(* IEC 61131-3 sources: plc-cip-batch-control/plc/prog, 5 files *)

(* ---- PRG_Alarms.st ---- *)
(*
    PRG_Alarms.st: the alarm list.

    Twelve points, each with a priority and an on-delay chosen so that the
    operator is not told about things that resolve themselves. ISA-18.2's first
    rule is that every alarm must require a response; a low chemical level that
    clears in two seconds does not.

    First-out is captured and held until the list goes quiet, so the record
    says which condition started the trip rather than which one is loudest by
    the time anyone looks.
*)

PROGRAM PRG_Alarms
VAR
    fbSafety        : FB_Alarm;
    fbSupplyPump    : FB_Alarm;
    fbReturnPump    : FB_Alarm;
    fbLevelLow      : FB_Alarm;
    fbCausticLow    : FB_Alarm;
    fbAcidLow       : FB_Alarm;
    fbTempLow       : FB_Alarm;
    fbFlowLow       : FB_Alarm;
    fbCircuitBusy   : FB_Alarm;
    fbPhaseTimeout  : FB_Alarm;
    fbNotClean      : FB_Alarm;
    fbNoSteam       : FB_Alarm;
    fbCondSensor    : FB_Alarm;
    i               : INT;
    xAnyLatched     : BOOL;
    xCirculating    : BOOL;
END_VAR

xCirculating := gxPhaseExecute AND (gPhaseStep = PS_CIRCULATE);

fbSafety(xCondition := gxSafetyTrip,
         iPriority  := 1,
         xAck       := xCmdAckAlarms,
         rNowS      := grPlcTimeS,
         stAlarm    := gAlarms[C_ALM_SAFETY]);

fbSupplyPump(xCondition := xSupplyPumpFault OR (xSupplyPumpRun AND NOT xSupplyPumpRunning),
             iPriority  := 1,
             tOnDelay   := T#5s,
             xAck       := xCmdAckAlarms,
             rNowS      := grPlcTimeS,
             stAlarm    := gAlarms[C_ALM_SUPPLY_PUMP]);

fbReturnPump(xCondition := xReturnPumpFault OR (xReturnPumpRun AND NOT xReturnPumpRunning),
             iPriority  := 2,
             tOnDelay   := T#5s,
             xAck       := xCmdAckAlarms,
             rNowS      := grPlcTimeS,
             stAlarm    := gAlarms[C_ALM_RETURN_PUMP]);

fbLevelLow(xCondition := (rLevelBalanceTankPct < C_LEVEL_TRIP_PCT) AND (gUnitState <> UST_IDLE),
           iPriority  := 2,
           tOnDelay   := T#3s,
           xAck       := xCmdAckAlarms,
           rNowS      := grPlcTimeS,
           stAlarm    := gAlarms[C_ALM_LEVEL_LOW]);

fbCausticLow(xCondition := rLevelCausticPct < C_CHEM_LEVEL_MIN,
             iPriority  := 3,
             tOnDelay   := T#10s,
             xAck       := xCmdAckAlarms,
             rNowS      := grPlcTimeS,
             stAlarm    := gAlarms[C_ALM_CAUSTIC_LOW]);

fbAcidLow(xCondition := rLevelAcidPct < C_CHEM_LEVEL_MIN,
          iPriority  := 3,
          tOnDelay   := T#10s,
          xAck       := xCmdAckAlarms,
          rNowS      := grPlcTimeS,
          stAlarm    := gAlarms[C_ALM_ACID_LOW]);

(* Twelve minutes: a cold circuit and a 1200 litre balance tank take about
   eight to come up to a wash temperature, so anything shorter alarms on every
   normal start. It still catches a steam valve that never opened. *)
fbTempLow(xCondition := xCirculating AND gPhaseParams.xHeat
                        AND (rTempReturnC < gPhaseParams.rTempMin),
          iPriority  := 2,
          tOnDelay   := T#12m,
          xAck       := xCmdAckAlarms,
          rNowS      := grPlcTimeS,
          stAlarm    := gAlarms[C_ALM_TEMP_LOW]);

fbFlowLow(xCondition := xCirculating AND (rFlowSupplyM3h < gPhaseParams.rFlowMin),
          iPriority  := 2,
          tOnDelay   := T#30s,
          xAck       := xCmdAckAlarms,
          rNowS      := grPlcTimeS,
          stAlarm    := gAlarms[C_ALM_FLOW_LOW]);

fbCircuitBusy(xCondition := (NOT xCircuitAvailable) AND (gUnitState <> UST_IDLE),
              iPriority  := 2,
              tOnDelay   := T#3s,
              xAck       := xCmdAckAlarms,
              rNowS      := grPlcTimeS,
              stAlarm    := gAlarms[C_ALM_CIRCUIT_BUSY]);

fbPhaseTimeout(xCondition := (gFailCode = FC_PHASE_TIMEOUT) OR (gFailCode = FC_CHARGE_TIMEOUT)
                             OR (gFailCode = FC_TEMP_TIMEOUT),
               iPriority  := 1,
               xAck       := xCmdAckAlarms,
               rNowS      := grPlcTimeS,
               stAlarm    := gAlarms[C_ALM_PHASE_TIMEOUT]);

fbNotClean(xCondition := gFailCode = FC_RINSE_NOT_CLEAN,
           iPriority  := 1,
           xAck       := xCmdAckAlarms,
           rNowS      := grPlcTimeS,
           stAlarm    := gAlarms[C_ALM_NOT_CLEAN]);

fbNoSteam(xCondition := (NOT xSteamAvailable) AND gPhaseParams.xHeat AND gxPhaseExecute,
          iPriority  := 3,
          tOnDelay   := T#10s,
          xAck       := xCmdAckAlarms,
          rNowS      := grPlcTimeS,
          stAlarm    := gAlarms[C_ALM_NO_STEAM]);

fbCondSensor(xCondition := gxCondSensorFault,
             iPriority  := 1,
             xAck       := xCmdAckAlarms,
             rNowS      := grPlcTimeS,
             stAlarm    := gAlarms[C_ALM_COND_SENSOR]);

(* ---- summary ---------------------------------------------------------- *)
giActiveAlarms := 0;
gxAlarmP1Active := FALSE;
xAnyLatched := FALSE;
xHmiAlarmHorn := FALSE;

FOR i := 1 TO C_ALARM_COUNT DO
    IF gAlarms[i].xLatched THEN
        xAnyLatched := TRUE;
        giActiveAlarms := giActiveAlarms + 1;
        IF gAlarms[i].xActive AND (gAlarms[i].iPriority = 1) THEN
            gxAlarmP1Active := TRUE;
        END_IF
        IF NOT gAlarms[i].xAcked THEN
            xHmiAlarmHorn := TRUE;
        END_IF
        IF giFirstOut = 0 THEN
            giFirstOut := i;
        END_IF
    END_IF
END_FOR

IF NOT xAnyLatched THEN
    giFirstOut := 0;
END_IF

(* Acknowledge is momentary too and this is the last program that reads it. *)
xCmdAckAlarms := FALSE;

END_PROGRAM

(* ---- PRG_Control.st ---- *)
(*
    PRG_Control.st: the only program that writes to the field outputs.

    It takes the demand PRG_Sequence produced, applies the permissives
    PRG_Safety produced and drives the valve matrix, the two motor starters
    and the two closed loops. Because it is the single writer, the question
    "what could possibly open the steam valve?" has exactly one answer.

    Loops:
      flow  -> supply pump speed, PI. Slow, because the pump is a VSD against
               a fixed circuit resistance and there is nothing to gain from
               being quick.
      temperature -> steam valve, PI on the supply temperature. Tuned soft:
               the plate pack has a couple of seconds of transport delay and
               the balance tank behind it is a 1200 litre integrator.
*)

PROGRAM PRG_Control
VAR
    fbFlowPid       : FB_Pid;
    fbTempPid       : FB_Pid;
    fbSupplyLimit   : FB_Pid;
    fbSupplyPump    : FB_Pump;
    fbReturnPump    : FB_Pump;
    xRunSupply      : BOOL;
    xRunReturn      : BOOL;
    xHeatDemand     : BOOL;
    xDoseDemand     : BOOL;
END_VAR

(* ---- interlocked demands --------------------------------------------- *)
xRunSupply  := gDemand.xSupplyPump AND gxPermitRun;
xRunReturn  := gDemand.xReturnPump AND gxPermitRun;
xHeatDemand := gDemand.xHeat AND gxPermitHeat;
xDoseDemand := gDemand.xDose AND gxPermitDose;

(* ---- motor starters --------------------------------------------------- *)
fbSupplyPump(xStart       := xRunSupply,
             xInterlockOk := gxPermitRun,
             xRunFeedback := xSupplyPumpRunning,
             xFault       := xSupplyPumpFault,
             xReset       := xCmdReset);

fbReturnPump(xStart       := xRunReturn,
             xInterlockOk := gxPermitRun,
             xRunFeedback := xReturnPumpRunning,
             xFault       := xReturnPumpFault,
             xReset       := xCmdReset);

xSupplyPumpRun := fbSupplyPump.xRun;
xReturnPumpRun := fbReturnPump.xRun;

(* ---- flow loop -------------------------------------------------------- *)
fbFlowPid(xEnable := fbSupplyPump.xRun,
          rPv     := rFlowSupplyM3h,
          rSp     := gDemand.rFlowSp,
          rKp     := 3.0,
          rTi     := 8.0,
          rOutMin := C_PUMP_SPEED_MIN,
          rOutMax := C_PUMP_SPEED_MAX,
          rCycleS := C_CYCLE_S);

IF fbSupplyPump.xRun THEN
    rSupplyPumpSpeedPct := fbFlowPid.rOut;
ELSE
    rSupplyPumpSpeedPct := 0.0;
END_IF

(* ---- temperature loop -------------------------------------------------- *)
(* The controlled variable is the return temperature, not the supply. The
   recipe specifies a temperature at the soil and the coldest point of the
   circuit is the one that has to reach it; controlling the supply instead
   throttles the steam as soon as one pass through the plate pack looks hot
   enough and the loop then takes three times as long to bring the balance
   tank up.

   Tuning is lambda tuning for an integrator with dead time: the circuit holds
   450 litres, so at 18 m3/h a change at the plate pack takes about 90 seconds
   to reach the return element. Kp 5 %/K, Ti 600 s. *)
fbTempPid(xEnable := xHeatDemand,
          rPv     := rTempReturnC,
          rSp     := gDemand.rTempSp,
          rKp     := 5.0,
          rTi     := 600.0,
          rOutMin := 0.0,
          rOutMax := 100.0,
          rCycleS := C_CYCLE_S);

(* Override: a proportional-only high limit on the plate-pack outlet, low
   selected against the main loop. Proportional only on purpose, because an
   integrator on the losing half of a selector winds up. *)
fbSupplyLimit(xEnable := xHeatDemand,
              rPv     := rTempSupplyC,
              rSp     := C_SUPPLY_TEMP_LIMIT,
              rKp     := 25.0,
              rTi     := 0.0,
              rOutMin := 0.0,
              rOutMax := 100.0,
              rCycleS := C_CYCLE_S);

xSteamIsolation := xHeatDemand;
IF xHeatDemand THEN
    rSteamValvePct := MIN(fbTempPid.rOut, fbSupplyLimit.rOut);
ELSE
    rSteamValvePct := 0.0;
END_IF

(* ---- valve matrix ----------------------------------------------------- *)
(* Source selection. Only one inlet is ever open and the fill valve gates
   the whole group so a phase can hold its line-up without taking liquid. *)
xV01FreshWater     := gDemand.xFillValve AND (gDemand.eSource = SRC_FRESH);
xV02RecoveredWater := gDemand.xFillValve AND (gDemand.eSource = SRC_RECOVERED);
xV11CausticSupply  := gDemand.xFillValve AND (gDemand.eSource = SRC_CAUSTIC);
xV12AcidSupply     := gDemand.xFillValve AND (gDemand.eSource = SRC_ACID);

(* Dosing is concentrate trim on top of whatever the tank already holds, so it
   is gated on the phase's dose demand rather than on the fill valve. *)
xV03CausticDose    := xDoseDemand AND (gDemand.eSource = SRC_CAUSTIC);
xV04AcidDose       := xDoseDemand AND (gDemand.eSource = SRC_ACID);

xV08ReturnToCaustic := FALSE;
xV10ReturnToAcid := FALSE;

(* Return destination. Exactly one of these is open whenever the return pump
   is running, so the circuit always has somewhere to discharge. *)
xV06ReturnToDrain    := FALSE;
xV07ReturnToBalance  := FALSE;
xV09ReturnToRecovery := FALSE;

CASE gDemand.eReturn OF
    RET_DRAIN:
        xV06ReturnToDrain := TRUE;
    RET_RECOVERY:
        xV09ReturnToRecovery := TRUE;
    RET_CAUSTIC:
        xV08ReturnToCaustic := TRUE;
    RET_ACID:
        xV10ReturnToAcid := TRUE;
    RET_BALANCE:
        xV07ReturnToBalance := TRUE;
END_CASE

xV05SupplyToCircuit := fbSupplyPump.xRun;

END_PROGRAM

(* ---- PRG_Kpi.st ---- *)
(*
    PRG_Kpi.st: consumption totals, the batch record and the SCADA image.

    Everything here is computed from instruments the skid actually has: the
    make-up flow meter, the supply flow meter, the two temperature elements
    either side of the heat exchanger and the dosing pump run time. Nothing
    is inferred from the model, so the same code would produce the same batch
    record on real hardware.

    Steam energy is the enthalpy the water gained across the plate pack:

        kW = m3/h * 1000 / 3600 [kg/s] * 4.19 [kJ/kg.K] * (Tsupply - Ttank) [K]

    which under-reports the boiler's fuel by the efficiency of the pack and
    the condensate return. It is the number the site can act on and it is
    the one the utility meter can be reconciled against.
*)

PROGRAM PRG_Kpi
VAR
    fbFresh         : FB_Totaliser;
    fbRecovered     : FB_Totaliser;
    fbEffluent      : FB_Totaliser;
    fbCaustic       : FB_Totaliser;
    fbAcid          : FB_Totaliser;
    fbEnergy        : FB_Totaliser;
    rEnergyKW       : REAL;
    rSnapWater      : REAL;
    rSnapChem       : REAL;
    rSnapEnergy     : REAL;
    i               : INT;
    xAllPass        : BOOL;
    xFinalRinseOk   : BOOL;
    xUnitActive     : BOOL;
END_VAR

xUnitActive := (gUnitState <> UST_IDLE)
               AND (gUnitState <> UST_COMPLETE)
               AND (gUnitState <> UST_ABORTED);

(* ---- instantaneous steam duty ---------------------------------------- *)
IF xSteamIsolation AND (rTempSupplyC > rTempBalanceTankC) THEN
    rEnergyKW := rFlowSupplyM3h * 1000.0 / 3600.0 * 4.19 * (rTempSupplyC - rTempBalanceTankC);
ELSE
    rEnergyKW := 0.0;
END_IF

(* ---- totalisers, all reset together at the start of a batch ------------
    Each is gated on the line-up rather than on a valve command. That
    distinction matters more than it looks.

    Make-up is bang-bang level control on a break tank, so V01 and V02 toggle
    every scan or two. The flow transmitter is read at the top of the scan and
    therefore reports the previous scan's flow, so gating the totaliser on the
    valve command aliases the two signals: on the scans the valve is open the
    meter is still reporting the scan it was shut, so the total comes out
    about a fifth low. The source selection only changes at a phase boundary
    and the meter reads zero when the valve is shut in any case. Gating on
    the source and letting the low-flow cut-off reject the noise measures
    what actually went through the meter.
*)
fbFresh(xEnable := gDemand.eSource = SRC_FRESH,
        rRatePerHour := rFlowMakeupM3h * 1000.0,
        rCutOff := 50.0,
        rCycleS := C_CYCLE_S,
        xReset := gxCycleReset);

fbRecovered(xEnable := gDemand.eSource = SRC_RECOVERED,
            rRatePerHour := rFlowMakeupM3h * 1000.0,
            rCutOff := 50.0,
            rCycleS := C_CYCLE_S,
            xReset := gxCycleReset);

fbEffluent(xEnable := xV06ReturnToDrain,
           rRatePerHour := rFlowSupplyM3h * 1000.0,
           rCutOff := 50.0,
           rCycleS := C_CYCLE_S,
           xReset := gxCycleReset);

fbCaustic(xEnable := xV03CausticDose,
          rRatePerHour := C_CAUSTIC_DOSE_LPM * 60.0,
          rCycleS := C_CYCLE_S,
          xReset := gxCycleReset);

fbAcid(xEnable := xV04AcidDose,
       rRatePerHour := C_ACID_DOSE_LPM * 60.0,
       rCycleS := C_CYCLE_S,
       xReset := gxCycleReset);

fbEnergy(xEnable := xSteamIsolation,
         rRatePerHour := rEnergyKW,
         rCycleS := C_CYCLE_S,
         xReset := gxCycleReset);

gKpi.rFreshWaterL     := fbFresh.rTotal;
gKpi.rRecoveredWaterL := fbRecovered.rTotal;
gKpi.rEffluentL       := fbEffluent.rTotal;
gKpi.rCausticL        := fbCaustic.rTotal;
gKpi.rAcidL           := fbAcid.rTotal;
gKpi.rEnergyKWh       := fbEnergy.rTotal;

IF gxCycleReset THEN
    grCycleElapsedS := 0.0;
    gKpi.xVerifiedClean := FALSE;
    rSnapWater := 0.0;
    rSnapChem := 0.0;
    rSnapEnergy := 0.0;
END_IF

IF xUnitActive THEN
    grCycleElapsedS := grCycleElapsedS + C_CYCLE_S;
END_IF
gKpi.rCycleTimeS := grCycleElapsedS;

(* ---- per-phase consumption, by difference ----------------------------- *)
IF gxPhaseStartPulse THEN
    rSnapWater  := fbFresh.rTotal + fbRecovered.rTotal;
    rSnapChem   := fbCaustic.rTotal + fbAcid.rTotal;
    rSnapEnergy := fbEnergy.rTotal;
END_IF

IF gxPhaseEndPulse AND (giPhaseIndex >= 1) AND (giPhaseIndex <= C_PHASE_COUNT) THEN
    gResults[giPhaseIndex].rWaterL := fbFresh.rTotal + fbRecovered.rTotal - rSnapWater;
    gResults[giPhaseIndex].rChemL := fbCaustic.rTotal + fbAcid.rTotal - rSnapChem;
    gResults[giPhaseIndex].rEnergyKWh := fbEnergy.rTotal - rSnapEnergy;
END_IF

(* ---- release criteria -------------------------------------------------- *)
(* A batch is only released if every phase that ran met its own criteria and
   the final rinse came back as clean as the water going in. A fixed-time
   recipe can complete without satisfying the second test and that is the
   whole argument for the adaptive one. *)
xAllPass := TRUE;
FOR i := 1 TO C_PHASE_COUNT DO
    IF gResults[i].xExecuted AND NOT gResults[i].xPass THEN
        xAllPass := FALSE;
    END_IF
END_FOR

xFinalRinseOk := gResults[5].xExecuted
                 AND gResults[5].xPass
                 AND (gResults[5].rEndConductivity <= gRecipe.rRinseEndCond);

IF gUnitState = UST_COMPLETE THEN
    gKpi.xVerifiedClean := xAllPass AND xFinalRinseOk;
END_IF

(* ---- SCADA image ------------------------------------------------------- *)
iHmiUnitState        := TO_INT(gUnitState);
iHmiPhase            := TO_INT(gPhase);
iHmiPhaseStep        := TO_INT(gPhaseStep);
iHmiFailCode         := TO_INT(gFailCode);
iHmiActiveAlarms     := giActiveAlarms;
iHmiFirstOutAlarm    := giFirstOut;
iHmiBatchId          := giBatchId;

rHmiFreshWaterL      := gKpi.rFreshWaterL;
rHmiRecoveredWaterL  := gKpi.rRecoveredWaterL;
rHmiEffluentL        := gKpi.rEffluentL;
rHmiCausticL         := gKpi.rCausticL;
rHmiAcidL            := gKpi.rAcidL;
rHmiEnergyKWh        := gKpi.rEnergyKWh;
rHmiCycleTimeS       := gKpi.rCycleTimeS;
rHmiPhaseElapsedS    := grPhaseElapsedS;
rHmiHoldAchievedS    := grHoldAchievedS;
rHmiConcentrationPct := grConcentrationPct;

xHmiVerifiedClean    := gKpi.xVerifiedClean;
xHmiCycleComplete    := gUnitState = UST_COMPLETE;
xHmiCycleAborted     := gUnitState = UST_ABORTED;
xHmiHeating          := xSteamIsolation;

END_PROGRAM

(* ---- PRG_Safety.st ---- *)
(*
    PRG_Safety.st: interlocks and permissives. First program in the task, so
    every other program sees a permit that was evaluated against this scan's
    inputs rather than the previous one's.

    Nothing here is a substitute for the hard-wired safety circuit. The E-stop
    drops the contactors and the steam solenoid directly; xSafetyOk is only the
    controller's view of that circuit, used to sequence a clean shutdown.

    Two interlocks earn their place:

      * no steam without proven flow. A steam-heated plate pack with no flow
        through it will boil the film against the plate, bake the soil on and
        eventually damage the gaskets.
      * no dosing without a running supply pump and a source that has stock in
        it, so concentrate cannot sit undiluted in the balance tank.
*)

PROGRAM PRG_Safety
VAR CONSTANT
    C_MIN_FLOW_HEAT : REAL := 8.0;      (* m3/h before steam may be admitted *)
    C_DRY_RUN_FLOW  : REAL := 2.0;      (* m3/h with the pump running is a dry run *)
END_VAR
VAR
    fbDryRun        : TON;
    fbCircuitLost   : TON;
    xChemStockOk    : BOOL;
END_VAR

grPlcTimeS := grPlcTimeS + C_CYCLE_S;

(* A running pump moving nothing is either dry or dead-headed. Either way it
   destroys the seal in minutes, so it is a latch-free hard stop. *)
fbDryRun(IN := xSupplyPumpRunning AND (rFlowSupplyM3h < C_DRY_RUN_FLOW), PT := T#20s);

fbCircuitLost(IN := NOT xCircuitAvailable, PT := T#3s);

gxSafetyTrip := (NOT xSafetyOk)
                OR xBalanceTankLowLow
                OR fbDryRun.Q
                OR (gUnitState <> UST_IDLE AND fbCircuitLost.Q);

gxPermitRun := xSafetyOk
               AND (NOT xBalanceTankLowLow)
               AND (NOT fbDryRun.Q)
               AND xCircuitAvailable
               AND (rLevelBalanceTankPct > C_LEVEL_TRIP_PCT);

gxPermitHeat := gxPermitRun
                AND xSteamAvailable
                AND xSupplyPumpRunning
                AND (rFlowSupplyM3h >= C_MIN_FLOW_HEAT);

(* Only the tank the current phase is drawing from has to have stock. *)
CASE gDemand.eSource OF
    SRC_CAUSTIC:
        xChemStockOk := rLevelCausticPct > C_CHEM_LEVEL_MIN;
    SRC_ACID:
        xChemStockOk := rLevelAcidPct > C_CHEM_LEVEL_MIN;
ELSE
    xChemStockOk := TRUE;
END_CASE

gxPermitDose := gxPermitRun AND xSupplyPumpRunning AND xChemStockOk;

END_PROGRAM

(* ---- PRG_Sequence.st ---- *)
(*
    PRG_Sequence.st: the ISA-88 unit procedure.

    This program owns the unit state machine and turns the recipe into phase
    parameters. It does not touch a single output. It produces a demand;
    PRG_Control decides whether the interlocks let that demand reach the
    field. Keeping the two apart is what makes the sequence readable and the
    interlocks auditable.

    Phase order is fixed; the recipe chooses which phases are in it:

        PRE_RINSE -> CAUSTIC -> INTERMEDIATE RINSE -> [ACID] ->
        FINAL RINSE -> [SANITISE] -> COMPLETE
*)

(*
    How long a rinse must run before its conductivity endpoint means anything.

    The return element sits downstream of the whole circuit, so a rinse that
    stops after twenty seconds has only measured the water that was already in
    the pipe. The floor is one and a half circuit turnovers at the recipe flow
    (135 seconds for a 450 litre circuit at 18 m3/h) or the recipe's own
    minimum, whichever is longer.
*)
FUNCTION RinseBlankTime : TIME
VAR_INPUT
    tFloor      : TIME;
    rFlowSpM3h  : REAL;
END_VAR
VAR
    rFlowLps    : REAL;
    rTurnoverS  : REAL;
END_VAR

rFlowLps := MAX(rFlowSpM3h, 1.0) * 1000.0 / 3600.0;
rTurnoverS := C_RINSE_TURNOVERS * C_CIRCUIT_VOLUME_L / rFlowLps;
RinseBlankTime := SecondsToTime(MAX(TimeToSeconds(tFloor), rTurnoverS));

END_FUNCTION

FUNCTION NextPhase : E_Phase
VAR_INPUT
    eCurrent     : E_Phase;
    xUseAcid     : BOOL;
    xUseSanitise : BOOL;
END_VAR

CASE eCurrent OF
    PH_IDLE:
        NextPhase := PH_PRE_RINSE;
    PH_PRE_RINSE:
        NextPhase := PH_CAUSTIC_WASH;
    PH_CAUSTIC_WASH:
        NextPhase := PH_INTERMEDIATE_RINSE;
    PH_INTERMEDIATE_RINSE:
        IF xUseAcid THEN
            NextPhase := PH_ACID_WASH;
        ELSE
            NextPhase := PH_FINAL_RINSE;
        END_IF
    PH_ACID_WASH:
        NextPhase := PH_FINAL_RINSE;
    PH_FINAL_RINSE:
        IF xUseSanitise THEN
            NextPhase := PH_SANITISE;
        ELSE
            NextPhase := PH_COMPLETE;
        END_IF
    PH_SANITISE:
        NextPhase := PH_COMPLETE;
ELSE
    NextPhase := PH_COMPLETE;
END_CASE

END_FUNCTION

PROGRAM PRG_Sequence
VAR
    fbUnit          : FB_UnitStateMachine;
    fbPhase         : FB_CipPhase;
    iPhaseIndex     : INT;
    iResultIndex    : INT;
    xReadyToStart   : BOOL;
    xProcComplete   : BOOL;
    xProcFailed     : BOOL;
    xPhaseGap       : BOOL;     (* one scan between phases, re-arms the engine *)
    xPhaseActive    : BOOL;     (* running or held: the engine keeps its state *)
    xExecutePhase   : BOOL;     (* running: accumulators and alarms advance *)
    ePrevPhase      : E_Phase;
END_VAR

(* ---------------------------------------------------------------------- *)
(* 1. Unit state machine                                                    *)
(* ---------------------------------------------------------------------- *)
xReadyToStart := (NOT gxSafetyTrip) AND xCircuitAvailable AND (NOT gxAlarmP1Active);

fbUnit(xStart              := xCmdStart,
       xHold               := xCmdHold,
       xRestart            := xCmdRestart,
       xAbort              := xCmdAbort,
       xReset              := xCmdReset,
       xReadyToStart       := xReadyToStart,
       xProcedureComplete  := xProcComplete,
       xProcedureFailed    := xProcFailed,
       xSafetyTrip         := gxSafetyTrip);

gUnitState := fbUnit.eState;

(* ---------------------------------------------------------------------- *)
(* 2. Start of batch                                                        *)
(* ---------------------------------------------------------------------- *)
gxCycleReset := FALSE;
IF fbUnit.xStartPulse THEN
    giBatchId := giBatchId + 1;
    gPhase := PH_PRE_RINSE;
    gFailCode := FC_NONE;
    xProcComplete := FALSE;
    xProcFailed := FALSE;
    xPhaseGap := FALSE;
    gxCycleReset := TRUE;
    gxCondSensorFault := FALSE;
    gxCondProven := FALSE;
    FOR iPhaseIndex := 1 TO C_PHASE_COUNT DO
        gResults[iPhaseIndex].ePhase := PH_IDLE;
        gResults[iPhaseIndex].xExecuted := FALSE;
        gResults[iPhaseIndex].xPass := FALSE;
        gResults[iPhaseIndex].eFail := FC_NONE;
        gResults[iPhaseIndex].rDurationS := 0.0;
        gResults[iPhaseIndex].rHoldAchievedS := 0.0;
        gResults[iPhaseIndex].rWaterL := 0.0;
        gResults[iPhaseIndex].rChemL := 0.0;
        gResults[iPhaseIndex].rEnergyKWh := 0.0;
    END_FOR
END_IF

IF fbUnit.eState = UST_IDLE THEN
    gPhase := PH_IDLE;
    gFailCode := FC_NONE;
END_IF

(* ---------------------------------------------------------------------- *)
(* 3. Phase parameters from the recipe                                      *)
(* ---------------------------------------------------------------------- *)
gPhaseParams.rFlowSp  := gRecipe.rFlowSp;
gPhaseParams.rFlowMin := gRecipe.rFlowMin;
gPhaseParams.tMaxPhase := gRecipe.tPhaseMax;
gPhaseParams.tMinPhase := T#30s;
gPhaseParams.xAdaptiveEnd := FALSE;
gPhaseParams.rEndConductivity := gRecipe.rRinseEndCond;
gPhaseParams.rConcSp := 0.0;
gPhaseParams.rConcMin := 0.0;
gPhaseParams.rConcMax := 0.0;
gPhaseParams.rTempSp := 0.0;
gPhaseParams.rTempMin := 0.0;
gPhaseParams.xHeat := FALSE;
gPhaseParams.xDose := FALSE;
gPhaseParams.xRecirculate := FALSE;

CASE gPhase OF

    PH_PRE_RINSE:
        (* Recovered final-rinse water if there is any, mains if not. This one
           line is most of the water saving: the pre-rinse is the biggest
           single-pass consumer in the cycle. *)
        IF rLevelRecoveryPct > 25.0 THEN
            gPhaseParams.eSource := SRC_RECOVERED;
        ELSE
            gPhaseParams.eSource := SRC_FRESH;
        END_IF
        gPhaseParams.eReturn := RET_DRAIN;
        gPhaseParams.tHold := gRecipe.tPreRinse;
        gPhaseParams.tMinPhase := RinseBlankTime(gRecipe.tRinseMin, gRecipe.rFlowSp);
        gPhaseParams.tRecover := T#20s;
        gPhaseParams.tMaxPhase := gRecipe.tRinseMax;
        gPhaseParams.xAdaptiveEnd := gRecipe.xAdaptive;
        (* Gross soil removal: a looser endpoint than the final rinse. *)
        gPhaseParams.rEndConductivity := gRecipe.rRinseEndCond * 3.0;

    PH_CAUSTIC_WASH:
        gPhaseParams.eSource := SRC_CAUSTIC;
        gPhaseParams.eReturn := RET_CAUSTIC;
        gPhaseParams.xRecirculate := TRUE;
        gPhaseParams.rTempSp := gRecipe.rCausticTempSp;
        gPhaseParams.rTempMin := gRecipe.rCausticTempMin;
        gPhaseParams.xHeat := TRUE;
        gPhaseParams.rConcSp := gRecipe.rCausticConcSp;
        gPhaseParams.rConcMin := gRecipe.rCausticConcSp - 0.25;
        gPhaseParams.rConcMax := gRecipe.rCausticConcSp + 0.50;
        gPhaseParams.xDose := TRUE;
        gPhaseParams.tHold := gRecipe.tCausticHold;
        gPhaseParams.tMinPhase := T#1m;
        gPhaseParams.tRecover := T#180s;

    PH_INTERMEDIATE_RINSE:
        gPhaseParams.eSource := SRC_FRESH;
        gPhaseParams.eReturn := RET_DRAIN;
        gPhaseParams.tHold := gRecipe.tIntRinse;
        gPhaseParams.tMinPhase := RinseBlankTime(gRecipe.tRinseMin, gRecipe.rFlowSp);
        gPhaseParams.tRecover := T#20s;
        gPhaseParams.tMaxPhase := gRecipe.tRinseMax;
        gPhaseParams.xAdaptiveEnd := gRecipe.xAdaptive;
        gPhaseParams.rEndConductivity := gRecipe.rRinseEndCond * 2.0;

    PH_ACID_WASH:
        gPhaseParams.eSource := SRC_ACID;
        gPhaseParams.eReturn := RET_ACID;
        gPhaseParams.xRecirculate := TRUE;
        gPhaseParams.rTempSp := gRecipe.rAcidTempSp;
        gPhaseParams.rTempMin := gRecipe.rAcidTempMin;
        gPhaseParams.xHeat := TRUE;
        gPhaseParams.rConcSp := gRecipe.rAcidConcSp;
        gPhaseParams.rConcMin := gRecipe.rAcidConcSp - 0.15;
        gPhaseParams.rConcMax := gRecipe.rAcidConcSp + 0.35;
        gPhaseParams.xDose := TRUE;
        gPhaseParams.tHold := gRecipe.tAcidHold;
        gPhaseParams.tMinPhase := T#1m;
        gPhaseParams.tRecover := T#180s;

    PH_FINAL_RINSE:
        gPhaseParams.eSource := SRC_FRESH;
        gPhaseParams.eReturn := RET_RECOVERY;
        gPhaseParams.tHold := gRecipe.tFinalRinse;
        gPhaseParams.tMinPhase := RinseBlankTime(gRecipe.tRinseMin, gRecipe.rFlowSp);
        gPhaseParams.tRecover := T#30s;
        gPhaseParams.tMaxPhase := gRecipe.tRinseMax;
        gPhaseParams.xAdaptiveEnd := gRecipe.xAdaptive;
        gPhaseParams.rEndConductivity := gRecipe.rRinseEndCond;

    PH_SANITISE:
        gPhaseParams.eSource := SRC_FRESH;
        gPhaseParams.eReturn := RET_BALANCE;
        gPhaseParams.xRecirculate := TRUE;
        gPhaseParams.rTempSp := gRecipe.rSanitiseTempSp;
        gPhaseParams.rTempMin := gRecipe.rSanitiseTempMin;
        gPhaseParams.xHeat := TRUE;
        gPhaseParams.tHold := gRecipe.tSanitiseHold;
        gPhaseParams.tMinPhase := T#1m;
        gPhaseParams.tRecover := T#30s;

ELSE
    gPhaseParams.eSource := SRC_NONE;
    gPhaseParams.eReturn := RET_DRAIN;
    gPhaseParams.tHold := T#0s;
    gPhaseParams.tRecover := T#0s;
END_CASE

(* ---------------------------------------------------------------------- *)
(* 3b. Derived measurements                                                 *)
(* ---------------------------------------------------------------------- *)
(* Both are computed here rather than in PRG_Control so the phase engine sees
   this scan's values instead of the previous scan's. The transmitter already
   compensates to 25 degC, so the calibration is a straight division. *)
grDeltaConductivity := rConductivityReturn - rConductivitySupply;

(* Strength is measured in the balance tank, not on the return line: during
   the charge step there is no established return flow to read. *)
CASE gPhaseParams.eSource OF
    SRC_CAUSTIC:
        grConcentrationPct := rConductivityTank / C_COND_K_CAUSTIC;
        grCondFloor := 0.5 * gPhaseParams.rConcSp * C_COND_K_CAUSTIC;
    SRC_ACID:
        grConcentrationPct := rConductivityTank / C_COND_K_ACID;
        grCondFloor := 0.5 * gPhaseParams.rConcSp * C_COND_K_ACID;
ELSE
    grConcentrationPct := 0.0;
    grCondFloor := 0.0;
END_CASE

(* ---------------------------------------------------------------------- *)
(* 4. Run the phase engine                                                  *)
(* ---------------------------------------------------------------------- *)
(* The engine stays executing through a hold so that it keeps its step, its
   elapsed time and its verified hold time. Dropping xExecute instead would
   look like the end of the phase and the restart would look like a fresh
   rising edge and begin the phase again from zero. *)
xPhaseActive := (fbUnit.xExecute OR fbUnit.xHolding)
                AND (gPhase <> PH_IDLE)
                AND (gPhase <> PH_COMPLETE)
                AND (NOT xPhaseGap);
xExecutePhase := xPhaseActive AND (NOT fbUnit.xHolding);

fbPhase(xExecute     := xPhaseActive,
        xHolding     := fbUnit.xHolding,
        ePhase       := gPhase,
        stParams     := gPhaseParams,
        rTempC       := rTempReturnC,
        rFlowM3h     := rFlowSupplyM3h,
        rConcPct     := grConcentrationPct,
        rDeltaCond   := grDeltaConductivity,
        rLevelPct    := rLevelBalanceTankPct,
        xPumpHealthy := NOT xSupplyPumpFault,
        rCycleS      := C_CYCLE_S);

gPhaseStep := fbPhase.eStep;
gDemand := fbPhase.stDemand;
grPhaseElapsedS := fbPhase.rElapsedS;
grHoldAchievedS := fbPhase.rHoldAchievedS;
gxPhaseExecute := xExecutePhase;
gxPhaseDone := fbPhase.xDone;
gxPhaseFailed := fbPhase.xFailed;

(*
    Plausibility check on the return conductivity element.

    Every rinse endpoint rests on this one transmitter; so does the
    release decision. The dangerous failure is not a dead reading but a
    reading stuck at something clean: an endpoint satisfied before the
    rinse began would pass a dirty circuit.

    There is one point in the cycle where the process guarantees a large
    signal. Circulating a wash at strength, the return line is full of
    detergent, so the element must at some point read at least half the
    expected value. A wash that finishes without it having done so means
    the element is not reading the process. Nothing may be released on its
    word.

    Written as a latch rather than a timer so that it holds for any hold
    time: a two minute wash proves the element as well as a twenty minute
    one. Both washes precede both rinses, so the check always runs before
    an endpoint is trusted.
*)
IF gxPhaseExecute
   AND (gPhaseStep = PS_CIRCULATE)
   AND (grCondFloor > 0.0)
   AND (rConductivityReturn >= grCondFloor) THEN
    gxCondProven := TRUE;
END_IF

(* ---------------------------------------------------------------------- *)
(* 5. Phase transitions and the batch record                                *)
(* ---------------------------------------------------------------------- *)
gxPhaseStartPulse := FALSE;
gxPhaseEndPulse := FALSE;
xPhaseGap := FALSE;

IF gPhase <> ePrevPhase THEN
    ePrevPhase := gPhase;
    IF (gPhase <> PH_IDLE) AND (gPhase <> PH_COMPLETE) THEN
        gxPhaseStartPulse := TRUE;
        gxCondProven := FALSE;
    END_IF
END_IF

iResultIndex := TO_INT(gPhase);

IF xExecutePhase AND fbPhase.xDone THEN
    gResults[iResultIndex] := fbPhase.stResult;
    gxPhaseEndPulse := TRUE;
    giPhaseIndex := iResultIndex;
    gPhase := NextPhase(gPhase, gRecipe.xUseAcid, gRecipe.xUseSanitise);
    xPhaseGap := TRUE;
END_IF

IF gxPhaseEndPulse AND (grCondFloor > 0.0) AND (NOT gxCondProven) THEN
    gxCondSensorFault := TRUE;
END_IF

IF gxCondSensorFault AND (gFailCode = FC_NONE) THEN
    gFailCode := FC_SENSOR_FAULT;
    xProcFailed := TRUE;
END_IF

IF xExecutePhase AND fbPhase.xFailed THEN
    gResults[iResultIndex] := fbPhase.stResult;
    gxPhaseEndPulse := TRUE;
    giPhaseIndex := iResultIndex;
    gFailCode := fbPhase.eFail;
    xProcFailed := TRUE;
END_IF

IF (gPhase = PH_COMPLETE) AND (fbUnit.eState = UST_RUNNING) THEN
    xProcComplete := TRUE;
END_IF

IF fbUnit.xAborting AND (gFailCode = FC_NONE) THEN
    IF gxSafetyTrip THEN
        gFailCode := FC_SAFETY_TRIP;
    ELSE
        gFailCode := FC_OPERATOR_ABORT;
    END_IF
END_IF

IF fbUnit.eState = UST_ABORTED THEN
    xProcFailed := FALSE;    (* consumed; the state machine is already there *)
END_IF

(* Momentary commands. The edges were taken at the top of this program, so the
   bits are cleared here and a client only ever has to set one. *)
xCmdStart := FALSE;
xCmdHold := FALSE;
xCmdRestart := FALSE;
xCmdAbort := FALSE;
xCmdReset := FALSE;

END_PROGRAM
